FUNCTION FC 1 : VOID
BEGIN
NETWORK
      L 40000
END_FUNCTION
